Universal Robots PolyScope program: TgtProg.urp

Program TgtProg (createdIn=3.0.0 lastSavedIn=3.0.0 directory=/programs installation=default)
Robot Program (runOnlyOnce=true motionType=MoveJ speed=1.047198 acceleration=1.396263 useActiveTCP=false)
  'Program generated by RoboDK v6.0.7 for UR10 on XX/XX/XXXX 18:00:00'
  'Using nominal kinematics.'
  Wait Sleep waitTime=0
  Wait Sleep waitTime=0.001
  Popup Message (haltProgram=false message=a <b> & "c" )
  'x <y> & 'z''
  MoveL speed 5 mm/s, acceleration 15000 mm/s^2 (useActiveTCP=true)
    Waypoint Waypoint_1: TCP in base x=-640 y=500 z=370 mm, rx=0.732 ry=2.1859 rz=-0.5703 rad; joints [0, -10, 20, 0, 30, 0] deg
  Script: movej([0.174533, -0.174533, 0.349066, 0.000000, 0.523599, 0.087266],39.99946,0.75000,0,0.0000)
  MoveJ speed 42.97 deg/s, acceleration 2291.77 deg/s^2 (useActiveTCP=true)
    Waypoint Waypoint_2: TCP in base x=-640 y=500 z=370 mm, rx=0.732 ry=2.1859 rz=-0.5703 rad; joints [10, -10, 20, 0, 30, 5] deg
